(* IEC 61131-3 sources: kns-port-domestic/tools/inventory_tests/fixtures/lib/src/DUTs, 5 files *)

(* ---- E_Mode.dut.st ---- *)
{attribute 'qualified_only'}
{attribute 'strict'}
// Режим устройства: перечисление с базовым типом
TYPE E_Mode :
(
    Auto := 0,
    Manual := 1
) INT;
END_TYPE

(* ---- ST_Base.dut.st ---- *)
// Базовая структура конфигурации
TYPE ST_Base :
STRUCT
    iLimit : INT;
END_STRUCT
END_TYPE

(* ---- ST_Ext.dut.st ---- *)
// Наследник структуры: 64-битные и широкие строки, поддиапазон
TYPE ST_Ext EXTENDS ST_Base :
STRUCT
    lwMask : LWORD;
    wsText : WSTRING(40);
    iPct : INT(0..100);
END_STRUCT
END_TYPE

(* ---- T_Percent.dut.st ---- *)
// Процент как псевдоним с поддиапазоном
TYPE T_Percent : INT(0..100);
END_TYPE

(* ---- U_Raw.dut.st ---- *)
// Сырое значение регистра
TYPE U_Raw :
UNION
    dwRaw : DWORD;
    rValue : REAL;
END_UNION
END_TYPE
